// TIA Portal V21 export
// export: Created 2026-11-10T07:35:06.5808748Z, ExportSetting WithDefaults, DisplayName Totally Integrated Automation Portal, DisplayVersion V21 Update 3, DisplayName STEP 7 Professional, DisplayVersion V21 Update 3, DisplayName STEP 7 Safety, DisplayVersion V21, DisplayName Tech WebApplication, DisplayVersion V21, DisplayName WinCC Basic/Comfort/Advanced, DisplayVersion V21 Update 3, DisplayName WinCC Unified, DisplayVersion V21 Update 3
FUNCTION_BLOCK "FB_Lad_ex050"   // FB95, LAD
{ S7_Optimized_Access := 'TRUE' }
VERSION : 0.1
// stored: AutoNumber true, IsIECCheckEnabled false, IsRetainMemResEnabled false, MemoryReserve 100, SetENOAutomatically false, UDAEnableTagReadback false
   VAR_INPUT
      v_id : HW_SUBMODULE;
      v_offset : Int;
      v_len : Int;
   END_VAR
   VAR_OUTPUT
      v_status : DWord;
      v_error : Bool;
   END_VAR
   VAR_IN_OUT
      v_outputs : Array[0..99] of Byte;
   END_VAR
   VAR
      inst { S7_SetPoint := 'True'} : SETIO_PART;
   END_VAR
BEGIN

REGION Network 1: SETIO_PART - Write outputs of a submodule
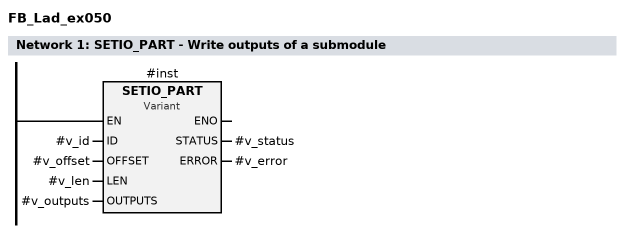
   RUNG wire#powerrail
      { S7_Templates := "[ptr_type := Variant, id_type := HW_SUBMODULE]" } #inst.SETIO_PART(ID := #v_id, OFFSET := #v_offset, LEN := #v_len, STATUS => #v_status, ERROR => #v_error, OUTPUTS := #v_outputs)
   END_RUNG
   // the same network as SCL:
   #inst(ID := #v_id,   // SETIO_PART
         OFFSET := #v_offset,
         LEN := #v_len,
         OUTPUTS := #v_outputs,
         STATUS => #v_status,
         ERROR => #v_error);
END_REGION
END_FUNCTION_BLOCK
